Fanuc KAREL source: KC00049.KL

PROGRAM KC00049
%NOLOCKGROUP
%ENVIRONMENT REGOPE
VAR
  I: INTEGER
  J: INTEGER
  K: INTEGER
  R: REAL
  B: BOOLEAN
  S: STRING[80]
  T: STRING[80]
  P: PATH
  Q: PATH
  AI: ARRAY[8] OF INTEGER
  AB: ARRAY[244] OF BYTE
  JP: JOINTPOS
BEGIN
  SET_TPE_JPOS_REG(I,JP,J)
END KC00049
